// TIA Portal V20 export
// export: Created 2026-10-19T18:03:04.8677323Z, ExportSetting WithDefaults, DisplayName Totally Integrated Automation Portal, DisplayVersion V20 Update 6, DisplayName TIA Portal Openness, DisplayVersion V20 Update 6, DisplayName TIA Portal Version Control Interface, DisplayVersion V20 Update 6, DisplayName SINAMICS Startdrive Advanced, DisplayVersion V20 SP1, DisplayName SINAMICS Startdrive G130, G150, S120, S150, SINAMICS MV, G220, S200, S210, DisplayVersion V20 SP1, DisplayName SINAMICS Startdrive G110M, G120, G120C, G120D, G120P, G115D, DisplayVersion V20 SP1, DisplayName STEP 7 Professional, DisplayVersion V20 Update 6, DisplayName STEP 7 Safety, DisplayVersion V20 Update 2, DisplayName WinCC Basic/Comfort/Advanced, DisplayVersion V20 Update 6, DisplayName WinCC Unified, DisplayVersion V20 Update 6
DATA_BLOCK "Stack_Lights_DB"   // DB62
VERSION : 0.1
// stored: AutoNumber true, DBAccessibleFromOPCUA true, DBAccessibleFromWebserver true, InstanceOfName Stack_Lights, InstanceOfType FB
"Stack_Lights"
   // VAR_INPUT
   //    VTD_Mode : UInt;
   //    Fault : Bool;
   // END_VAR
   // VAR_OUTPUT
   //    Red : Bool;
   //    Green : Bool;
   //    Blue : Bool;
   //    Buzzer : Bool;
   // END_VAR
BEGIN
END_DATA_BLOCK
